// TIA Portal V20 export
// export: Created 2026-10-06T00:00:00
Screen "Start"  1280x800, Number=1, Template=Base
  ScreenLayer 
    Rectangle "Logo" at 20,100 size 40x40
